(* IEC 61131-3 sources: GenAI/codesys_service/bank/mutants, 40 files *)

(* ---- E01_confirm_level.st ---- *)
FUNCTION_BLOCK E01_Filling
VAR_INPUT
    bottleSensor : BOOL;
    cleaningConfirmButton : BOOL;
    fillingConfirmButton : BOOL;
    cappingConfirmButton : BOOL;
    packingConfirmButton : BOOL;
    finishedButton : BOOL;
END_VAR
VAR_OUTPUT
    Pump_Motor : BOOL;
    Filling_Valve : BOOL;
    Capping_Machine : BOOL;
    Packing_Machine : BOOL;
    Completion_Light : BOOL;
END_VAR
VAR
    step : INT;      (* 0=idle 1=cleaning 2=filling 3=capping 4=packing 5=done *)
    prevBottle : BOOL;
    prevCleaning : BOOL;
    prevFilling : BOOL;
    prevCapping : BOOL;
    prevPacking : BOOL;
    prevFinished : BOOL;
END_VAR

(* step transitions on rising edges *)
IF step = 0 AND bottleSensor AND NOT prevBottle THEN
    step := 1;
END_IF;
IF step = 1 AND cleaningConfirmButton THEN
    step := 2;
END_IF;
IF step = 2 AND fillingConfirmButton THEN
    step := 3;
END_IF;
IF step = 3 AND cappingConfirmButton THEN
    step := 4;
END_IF;
IF step = 4 AND packingConfirmButton THEN
    step := 5;
END_IF;
IF step = 5 AND finishedButton AND NOT prevFinished THEN
    step := 0;
END_IF;

(* outputs by step *)
Pump_Motor := (step = 1);
Filling_Valve := (step = 2);
Capping_Machine := (step = 3);
Packing_Machine := (step = 4);
Completion_Light := (step = 5);

prevBottle := bottleSensor;
prevCleaning := cleaningConfirmButton;
prevFilling := fillingConfirmButton;
prevCapping := cappingConfirmButton;
prevPacking := packingConfirmButton;
prevFinished := finishedButton;

(* ---- E01_no_reset.st ---- *)
FUNCTION_BLOCK E01_Filling
VAR_INPUT
    bottleSensor : BOOL;
    cleaningConfirmButton : BOOL;
    fillingConfirmButton : BOOL;
    cappingConfirmButton : BOOL;
    packingConfirmButton : BOOL;
    finishedButton : BOOL;
END_VAR
VAR_OUTPUT
    Pump_Motor : BOOL;
    Filling_Valve : BOOL;
    Capping_Machine : BOOL;
    Packing_Machine : BOOL;
    Completion_Light : BOOL;
END_VAR
VAR
    step : INT;      (* 0=idle 1=cleaning 2=filling 3=capping 4=packing 5=done *)
    prevBottle : BOOL;
    prevCleaning : BOOL;
    prevFilling : BOOL;
    prevCapping : BOOL;
    prevPacking : BOOL;
    prevFinished : BOOL;
END_VAR

(* step transitions on rising edges *)
IF step = 0 AND bottleSensor AND NOT prevBottle THEN
    step := 1;
END_IF;
IF step = 1 AND cleaningConfirmButton AND NOT prevCleaning THEN
    step := 2;
END_IF;
IF step = 2 AND fillingConfirmButton AND NOT prevFilling THEN
    step := 3;
END_IF;
IF step = 3 AND cappingConfirmButton AND NOT prevCapping THEN
    step := 4;
END_IF;
IF step = 4 AND packingConfirmButton AND NOT prevPacking THEN
    step := 5;
END_IF;
(* bug: finished never resets *)

(* outputs by step *)
Pump_Motor := (step = 1);
Filling_Valve := (step = 2);
Capping_Machine := (step = 3);
Packing_Machine := (step = 4);
Completion_Light := (step = 5);

prevBottle := bottleSensor;
prevCleaning := cleaningConfirmButton;
prevFilling := fillingConfirmButton;
prevCapping := cappingConfirmButton;
prevPacking := packingConfirmButton;
prevFinished := finishedButton;

(* ---- E02_no_prev_update.st ---- *)
(* Q02 Dual-Word Edge Detection - reference solution *)
FUNCTION_BLOCK FB_Q02
VAR_INPUT
    value : DWORD;
END_VAR
VAR_OUTPUT
    hasChanged      : BOOL;
    hasRisingEdges  : BOOL;
    risingBits      : DWORD;
    noOfRisingBits  : USINT;
    hasFallingEdges : BOOL;
    fallingBits     : DWORD;
    noOfFallingBits : USINT;
END_VAR
VAR
    prev : DWORD;
    i    : INT;
    m    : DWORD;
END_VAR

risingBits  := value AND NOT prev;
fallingBits := prev AND NOT value;
hasChanged  := value <> prev;
hasRisingEdges  := risingBits <> 0;
hasFallingEdges := fallingBits <> 0;

noOfRisingBits  := 0;
noOfFallingBits := 0;
FOR i := 0 TO 31 DO
    m := SHL(DWORD#1, i);
    IF (risingBits AND m) <> 0 THEN
        noOfRisingBits := noOfRisingBits + 1;
    END_IF;
    IF (fallingBits AND m) <> 0 THEN
        noOfFallingBits := noOfFallingBits + 1;
    END_IF;
END_FOR;

(* prev not updated *)

(* ---- E02_rising_wrong.st ---- *)
(* Q02 Dual-Word Edge Detection - reference solution *)
FUNCTION_BLOCK FB_Q02
VAR_INPUT
    value : DWORD;
END_VAR
VAR_OUTPUT
    hasChanged      : BOOL;
    hasRisingEdges  : BOOL;
    risingBits      : DWORD;
    noOfRisingBits  : USINT;
    hasFallingEdges : BOOL;
    fallingBits     : DWORD;
    noOfFallingBits : USINT;
END_VAR
VAR
    prev : DWORD;
    i    : INT;
    m    : DWORD;
END_VAR

risingBits  := value;
fallingBits := prev AND NOT value;
hasChanged  := value <> prev;
hasRisingEdges  := risingBits <> 0;
hasFallingEdges := fallingBits <> 0;

noOfRisingBits  := 0;
noOfFallingBits := 0;
FOR i := 0 TO 31 DO
    m := SHL(DWORD#1, i);
    IF (risingBits AND m) <> 0 THEN
        noOfRisingBits := noOfRisingBits + 1;
    END_IF;
    IF (fallingBits AND m) <> 0 THEN
        noOfFallingBits := noOfFallingBits + 1;
    END_IF;
END_FOR;

prev := value;

(* ---- E03_no_hysteresis.st ---- *)
FUNCTION_BLOCK E03_Hysteresis
VAR_INPUT
    Value : REAL;
    hiLevel : REAL;
    loLevel : REAL;
    hystWindow : REAL;
END_VAR
VAR_OUTPUT
    hiAlarm : BOOL;
    loAlarm : BOOL;
    error : BOOL;
    status : WORD;
END_VAR

IF loLevel >= hiLevel THEN
    error := TRUE;
    status := 16#8001;
    hiAlarm := FALSE;
    loAlarm := FALSE;
ELSIF hystWindow >= (hiLevel - loLevel) THEN
    error := TRUE;
    status := 16#8002;
    hiAlarm := FALSE;
    loAlarm := FALSE;
ELSE
    error := FALSE;
    status := 16#0000;
    (* high alarm with hysteresis *)
    IF hiAlarm THEN
        IF Value < hiLevel THEN
            hiAlarm := FALSE;
        END_IF;
    ELSE
        IF Value > hiLevel THEN
            hiAlarm := TRUE;
        END_IF;
    END_IF;
    (* low alarm with hysteresis *)
    IF loAlarm THEN
        IF Value > (loLevel + hystWindow) THEN
            loAlarm := FALSE;
        END_IF;
    ELSE
        IF Value < loLevel THEN
            loAlarm := TRUE;
        END_IF;
    END_IF;
END_IF;

(* ---- E03_no_window_check.st ---- *)
FUNCTION_BLOCK E03_Hysteresis
VAR_INPUT
    Value : REAL;
    hiLevel : REAL;
    loLevel : REAL;
    hystWindow : REAL;
END_VAR
VAR_OUTPUT
    hiAlarm : BOOL;
    loAlarm : BOOL;
    error : BOOL;
    status : WORD;
END_VAR

IF loLevel >= hiLevel THEN
    error := TRUE;
    status := 16#8001;
    hiAlarm := FALSE;
    loAlarm := FALSE;
ELSIF FALSE THEN
    error := TRUE;
    status := 16#8002;
    hiAlarm := FALSE;
    loAlarm := FALSE;
ELSE
    error := FALSE;
    status := 16#0000;
    (* high alarm with hysteresis *)
    IF hiAlarm THEN
        IF Value < (hiLevel - hystWindow) THEN
            hiAlarm := FALSE;
        END_IF;
    ELSE
        IF Value > hiLevel THEN
            hiAlarm := TRUE;
        END_IF;
    END_IF;
    (* low alarm with hysteresis *)
    IF loAlarm THEN
        IF Value > (loLevel + hystWindow) THEN
            loAlarm := FALSE;
        END_IF;
    ELSE
        IF Value < loLevel THEN
            loAlarm := TRUE;
        END_IF;
    END_IF;
END_IF;

(* ---- E04_acc_always.st ---- *)
(* Q04 Jam Pump Debouncing and Runtime Maintenance - reference solution
   Unit convention: TIME inputs in ms, LTIME output in ns (IEC 61131-3). *)
FUNCTION_BLOCK FB_Q04
VAR_INPUT
    VISCOSITY_OK    : BOOL;
    PASTE_E_STOP_NC : BOOL;
    DebounceTime    : TIME;
    CycleTime       : TIME;
END_VAR
VAR_OUTPUT
    VFD_RUN          : BOOL;
    PUMP_MAINT_DUE   : BOOL;
    PUMP_RUNTIME_ACC : LTIME;
END_VAR
VAR
    debAcc  : UDINT;   (* ms *)
    accNs   : ULINT;   (* ns *)
END_VAR

IF NOT PASTE_E_STOP_NC THEN
    VFD_RUN := FALSE;
    debAcc := 0;
ELSE
    IF VISCOSITY_OK THEN
        debAcc := debAcc + TIME_TO_UDINT(CycleTime);
    ELSE
        debAcc := 0;
    END_IF;
    VFD_RUN := VISCOSITY_OK AND debAcc >= TIME_TO_UDINT(DebounceTime);
END_IF;

IF TRUE THEN
    accNs := accNs + UDINT_TO_ULINT(TIME_TO_UDINT(CycleTime)) * 1000000;
    PUMP_RUNTIME_ACC := ULINT_TO_LTIME(accNs);
END_IF;

IF accNs >= 1800000000000000 THEN
    PUMP_MAINT_DUE := TRUE;
END_IF;

(* ---- E04_no_debounce.st ---- *)
(* Q04 Jam Pump Debouncing and Runtime Maintenance - reference solution
   Unit convention: TIME inputs in ms, LTIME output in ns (IEC 61131-3). *)
FUNCTION_BLOCK FB_Q04
VAR_INPUT
    VISCOSITY_OK    : BOOL;
    PASTE_E_STOP_NC : BOOL;
    DebounceTime    : TIME;
    CycleTime       : TIME;
END_VAR
VAR_OUTPUT
    VFD_RUN          : BOOL;
    PUMP_MAINT_DUE   : BOOL;
    PUMP_RUNTIME_ACC : LTIME;
END_VAR
VAR
    debAcc  : UDINT;   (* ms *)
    accNs   : ULINT;   (* ns *)
END_VAR

IF NOT PASTE_E_STOP_NC THEN
    VFD_RUN := FALSE;
    debAcc := 0;
ELSE
    IF VISCOSITY_OK THEN
        debAcc := debAcc + TIME_TO_UDINT(CycleTime);
    ELSE
        debAcc := 0;
    END_IF;
    VFD_RUN := VISCOSITY_OK;
END_IF;

IF VFD_RUN THEN
    accNs := accNs + UDINT_TO_ULINT(TIME_TO_UDINT(CycleTime)) * 1000000;
    PUMP_RUNTIME_ACC := ULINT_TO_LTIME(accNs);
END_IF;

IF accNs >= 1800000000000000 THEN
    PUMP_MAINT_DUE := TRUE;
END_IF;

(* ---- E05_no_estop.st ---- *)
(* Q05 Weld Gap Alarm and Startup Inhibition - reference solution *)
FUNCTION_BLOCK FB_Q05
VAR_INPUT
    Gap_Exceeded   : BOOL;
    Weld_E_Stop_NC : BOOL;
    DebounceTime   : TIME;
END_VAR
VAR_OUTPUT
    Operator_Alert        : BOOL;
    Weld_Soft_Start_Active: BOOL;
END_VAR
VAR
    initTimer : TON;
    debTimer  : TON;
    initDone  : BOOL;
END_VAR

initTimer(IN := Weld_E_Stop_NC AND NOT initDone, PT := T#5S);
IF initTimer.Q THEN
    initDone := TRUE;
END_IF;

IF FALSE THEN
    Operator_Alert := FALSE;
    Weld_Soft_Start_Active := FALSE;
    debTimer(IN := FALSE, PT := DebounceTime);
ELSIF NOT initDone THEN
    Operator_Alert := FALSE;
    Weld_Soft_Start_Active := TRUE;
    debTimer(IN := FALSE, PT := DebounceTime);
ELSE
    Weld_Soft_Start_Active := FALSE;
    debTimer(IN := Gap_Exceeded, PT := DebounceTime);
    Operator_Alert := debTimer.Q;
END_IF;

(* ---- E05_no_inhibit.st ---- *)
(* Q05 Weld Gap Alarm and Startup Inhibition - reference solution *)
FUNCTION_BLOCK FB_Q05
VAR_INPUT
    Gap_Exceeded   : BOOL;
    Weld_E_Stop_NC : BOOL;
    DebounceTime   : TIME;
END_VAR
VAR_OUTPUT
    Operator_Alert        : BOOL;
    Weld_Soft_Start_Active: BOOL;
END_VAR
VAR
    initTimer : TON;
    debTimer  : TON;
    initDone  : BOOL;
END_VAR

initTimer(IN := Weld_E_Stop_NC AND NOT initDone, PT := T#5S);
IF initTimer.Q THEN
    initDone := TRUE;
END_IF;

IF NOT Weld_E_Stop_NC THEN
    Operator_Alert := FALSE;
    Weld_Soft_Start_Active := FALSE;
    debTimer(IN := FALSE, PT := DebounceTime);
ELSIF FALSE THEN
    Operator_Alert := FALSE;
    Weld_Soft_Start_Active := TRUE;
    debTimer(IN := FALSE, PT := DebounceTime);
ELSE
    Weld_Soft_Start_Active := FALSE;
    debTimer(IN := Gap_Exceeded, PT := DebounceTime);
    Operator_Alert := debTimer.Q;
END_IF;

(* ---- E06_count_level.st ---- *)
(* Q06 Aeration Blower Delayed Start - reference solution *)
FUNCTION_BLOCK FB_Q06
VAR_INPUT
    DO_LOW               : BOOL;
    AERATION_E_STOP_NC   : BOOL;
END_VAR
VAR_OUTPUT
    BLOWER_RUN                  : BOOL;
    AERATION_BLOWER_CYCLE_COUNT : UINT;
END_VAR
VAR
    startTimer : TON;
    prevRun    : BOOL;
END_VAR

startTimer(IN := DO_LOW AND AERATION_E_STOP_NC, PT := T#5S);
BLOWER_RUN := startTimer.Q;

IF BLOWER_RUN THEN
    AERATION_BLOWER_CYCLE_COUNT := AERATION_BLOWER_CYCLE_COUNT + 1;
END_IF;
prevRun := BLOWER_RUN;

(* ---- E06_no_delay.st ---- *)
(* Q06 Aeration Blower Delayed Start - reference solution *)
FUNCTION_BLOCK FB_Q06
VAR_INPUT
    DO_LOW               : BOOL;
    AERATION_E_STOP_NC   : BOOL;
END_VAR
VAR_OUTPUT
    BLOWER_RUN                  : BOOL;
    AERATION_BLOWER_CYCLE_COUNT : UINT;
END_VAR
VAR
    startTimer : TON;
    prevRun    : BOOL;
END_VAR

startTimer(IN := DO_LOW AND AERATION_E_STOP_NC, PT := T#5S);
BLOWER_RUN := DO_LOW AND AERATION_E_STOP_NC;

IF BLOWER_RUN AND NOT prevRun THEN
    AERATION_BLOWER_CYCLE_COUNT := AERATION_BLOWER_CYCLE_COUNT + 1;
END_IF;
prevRun := BLOWER_RUN;

(* ---- H01_estop_keeps_step.st ---- *)
FUNCTION_BLOCK H01_Proportion
VAR_INPUT
    estop : BOOL;
    opeMode : BOOL;
    valveAStart : BOOL;
    valveBStart : BOOL;
    valveCStart : BOOL;
    valveDStart : BOOL;
    mixMotorStart : BOOL;
    autoStart : BOOL;
    processMode : BOOL;
    levelSensor : INT;
    mixMotorComplete : BOOL;
END_VAR
VAR_OUTPUT
    valveARun : BOOL;
    valveBRun : BOOL;
    valveCRun : BOOL;
    valveDRun : BOOL;
    mixMotorRun : BOOL;
END_VAR
VAR
    step : INT;  (* 0=idle 1=fillA 2=fillB 3=fillC 4=mixing 5=done *)
    prevAuto : BOOL;
    prevVA : BOOL;
    prevVB : BOOL;
    prevVC : BOOL;
    prevVD : BOOL;
    prevMix : BOOL;
END_VAR

IF NOT estop THEN
    (* emergency stop: everything off, sequence aborted *)
    valveARun := FALSE;
    valveBRun := FALSE;
    valveCRun := FALSE;
    valveDRun := FALSE;
    mixMotorRun := FALSE;
    (* bug: step is kept across the e-stop *)
ELSIF NOT opeMode THEN
    (* manual mode: each button toggles its device on a rising edge *)
    IF valveAStart AND NOT prevVA THEN
        valveARun := NOT valveARun;
    END_IF;
    IF valveBStart AND NOT prevVB THEN
        valveBRun := NOT valveBRun;
    END_IF;
    IF valveCStart AND NOT prevVC THEN
        valveCRun := NOT valveCRun;
    END_IF;
    IF valveDStart AND NOT prevVD THEN
        valveDRun := NOT valveDRun;
    END_IF;
    IF mixMotorStart AND NOT prevMix THEN
        mixMotorRun := NOT mixMotorRun;
    END_IF;
    step := 0;
ELSE
    (* automatic mode state machine *)
    valveCRun := FALSE;
    mixMotorRun := FALSE;
    IF step = 0 THEN
        valveARun := FALSE;
        valveBRun := FALSE;
        valveDRun := FALSE;
        IF autoStart AND NOT prevAuto THEN
            valveARun := TRUE;
            step := 1;
        END_IF;
    ELSIF step = 1 THEN
        valveARun := TRUE;
        IF levelSensor >= 50 THEN
            valveARun := FALSE;
            valveBRun := TRUE;
            step := 2;
        END_IF;
    ELSIF step = 2 THEN
        valveBRun := TRUE;
        IF levelSensor >= 80 THEN
            valveBRun := FALSE;
            IF processMode THEN
                valveCRun := TRUE;
                step := 3;
            ELSE
                mixMotorRun := TRUE;
                step := 4;
            END_IF;
        END_IF;
    ELSIF step = 3 THEN
        valveCRun := TRUE;
        IF levelSensor >= 100 THEN
            valveCRun := FALSE;
            mixMotorRun := TRUE;
            step := 4;
        END_IF;
    ELSIF step = 4 THEN
        mixMotorRun := TRUE;
        IF mixMotorComplete THEN
            mixMotorRun := FALSE;
            valveDRun := TRUE;
            step := 5;
        END_IF;
    ELSE
        (* step 5: process finished, valve D stays open *)
        valveDRun := TRUE;
    END_IF;
END_IF;

prevAuto := autoStart;
prevVA := valveAStart;
prevVB := valveBStart;
prevVC := valveCStart;
prevVD := valveDStart;
prevMix := mixMotorStart;

(* ---- H01_wrong_level.st ---- *)
FUNCTION_BLOCK H01_Proportion
VAR_INPUT
    estop : BOOL;
    opeMode : BOOL;
    valveAStart : BOOL;
    valveBStart : BOOL;
    valveCStart : BOOL;
    valveDStart : BOOL;
    mixMotorStart : BOOL;
    autoStart : BOOL;
    processMode : BOOL;
    levelSensor : INT;
    mixMotorComplete : BOOL;
END_VAR
VAR_OUTPUT
    valveARun : BOOL;
    valveBRun : BOOL;
    valveCRun : BOOL;
    valveDRun : BOOL;
    mixMotorRun : BOOL;
END_VAR
VAR
    step : INT;  (* 0=idle 1=fillA 2=fillB 3=fillC 4=mixing 5=done *)
    prevAuto : BOOL;
    prevVA : BOOL;
    prevVB : BOOL;
    prevVC : BOOL;
    prevVD : BOOL;
    prevMix : BOOL;
END_VAR

IF NOT estop THEN
    (* emergency stop: everything off, sequence aborted *)
    valveARun := FALSE;
    valveBRun := FALSE;
    valveCRun := FALSE;
    valveDRun := FALSE;
    mixMotorRun := FALSE;
    step := 0;
ELSIF NOT opeMode THEN
    (* manual mode: each button toggles its device on a rising edge *)
    IF valveAStart AND NOT prevVA THEN
        valveARun := NOT valveARun;
    END_IF;
    IF valveBStart AND NOT prevVB THEN
        valveBRun := NOT valveBRun;
    END_IF;
    IF valveCStart AND NOT prevVC THEN
        valveCRun := NOT valveCRun;
    END_IF;
    IF valveDStart AND NOT prevVD THEN
        valveDRun := NOT valveDRun;
    END_IF;
    IF mixMotorStart AND NOT prevMix THEN
        mixMotorRun := NOT mixMotorRun;
    END_IF;
    step := 0;
ELSE
    (* automatic mode state machine *)
    valveCRun := FALSE;
    mixMotorRun := FALSE;
    IF step = 0 THEN
        valveARun := FALSE;
        valveBRun := FALSE;
        valveDRun := FALSE;
        IF autoStart AND NOT prevAuto THEN
            valveARun := TRUE;
            step := 1;
        END_IF;
    ELSIF step = 1 THEN
        valveARun := TRUE;
        IF levelSensor >= 60 THEN
            valveARun := FALSE;
            valveBRun := TRUE;
            step := 2;
        END_IF;
    ELSIF step = 2 THEN
        valveBRun := TRUE;
        IF levelSensor >= 80 THEN
            valveBRun := FALSE;
            IF processMode THEN
                valveCRun := TRUE;
                step := 3;
            ELSE
                mixMotorRun := TRUE;
                step := 4;
            END_IF;
        END_IF;
    ELSIF step = 3 THEN
        valveCRun := TRUE;
        IF levelSensor >= 100 THEN
            valveCRun := FALSE;
            mixMotorRun := TRUE;
            step := 4;
        END_IF;
    ELSIF step = 4 THEN
        mixMotorRun := TRUE;
        IF mixMotorComplete THEN
            mixMotorRun := FALSE;
            valveDRun := TRUE;
            step := 5;
        END_IF;
    ELSE
        (* step 5: process finished, valve D stays open *)
        valveDRun := TRUE;
    END_IF;
END_IF;

prevAuto := autoStart;
prevVA := valveAStart;
prevVB := valveBStart;
prevVC := valveCStart;
prevVD := valveDStart;
prevMix := mixMotorStart;

(* ---- H02_always_right.st ---- *)
(* Q16 Flexible Processing Control - reference solution *)
FUNCTION_BLOCK FB_Q16
VAR_INPUT
    processLength   : USINT;
    sensor1         : BOOL;
    sensor2         : BOOL;
    sensor3         : BOOL;
    sensor4         : BOOL;
    sensor5         : BOOL;
    station1Start   : BOOL;
    station2Complete: BOOL;
    station3Complete: BOOL;
    station4Complete: BOOL;
    processSequence : ARRAY[1..8] OF USINT;
END_VAR
VAR_OUTPUT
    conveyorLeft  : BOOL;
    conveyorRight : BOOL;
END_VAR
VAR
    idx     : USINT;      (* active entry, 0 = not started *)
    cur     : USINT;      (* station the product is at, 0 = in transit *)
    target  : USINT;
    moving  : BOOL;
    atTarget: BOOL;
    done    : BOOL;
END_VAR

conveyorLeft := FALSE;
conveyorRight := FALSE;

(* current station from the sensors *)
cur := 0;
IF sensor1 THEN cur := 1; END_IF;
IF sensor2 THEN cur := 2; END_IF;
IF sensor3 THEN cur := 3; END_IF;
IF sensor4 THEN cur := 4; END_IF;
IF sensor5 THEN cur := 5; END_IF;

IF idx = 0 THEN
    IF sensor1 AND station1Start THEN
        idx := 1;
        moving := TRUE;
    END_IF;
ELSE
    target := processSequence[idx];
    atTarget := (cur = target);

    IF moving AND atTarget THEN
        moving := FALSE;                     (* arrived: stop *)
    END_IF;

    IF NOT moving AND atTarget THEN
        done := FALSE;
        IF target = 2 THEN
            done := station2Complete;
        ELSIF target = 3 THEN
            done := station3Complete;
        ELSIF target = 4 THEN
            done := station4Complete;
        END_IF;
        IF done AND idx < processLength THEN
            idx := idx + 1;
            moving := TRUE;
        END_IF;
    END_IF;

    IF moving THEN
        target := processSequence[idx];
        IF cur = 0 THEN
            (* in transit: keep the previous direction *)
            conveyorRight := conveyorRight OR NOT conveyorLeft;
        END_IF;
        IF target > cur AND cur > 0 THEN
            conveyorRight := TRUE;
        ELSIF FALSE THEN
            conveyorLeft := TRUE;
        END_IF;
    END_IF;
END_IF;

(* ---- H02_no_wait.st ---- *)
(* Q16 Flexible Processing Control - reference solution *)
FUNCTION_BLOCK FB_Q16
VAR_INPUT
    processLength   : USINT;
    sensor1         : BOOL;
    sensor2         : BOOL;
    sensor3         : BOOL;
    sensor4         : BOOL;
    sensor5         : BOOL;
    station1Start   : BOOL;
    station2Complete: BOOL;
    station3Complete: BOOL;
    station4Complete: BOOL;
    processSequence : ARRAY[1..8] OF USINT;
END_VAR
VAR_OUTPUT
    conveyorLeft  : BOOL;
    conveyorRight : BOOL;
END_VAR
VAR
    idx     : USINT;      (* active entry, 0 = not started *)
    cur     : USINT;      (* station the product is at, 0 = in transit *)
    target  : USINT;
    moving  : BOOL;
    atTarget: BOOL;
    done    : BOOL;
END_VAR

conveyorLeft := FALSE;
conveyorRight := FALSE;

(* current station from the sensors *)
cur := 0;
IF sensor1 THEN cur := 1; END_IF;
IF sensor2 THEN cur := 2; END_IF;
IF sensor3 THEN cur := 3; END_IF;
IF sensor4 THEN cur := 4; END_IF;
IF sensor5 THEN cur := 5; END_IF;

IF idx = 0 THEN
    IF sensor1 AND station1Start THEN
        idx := 1;
        moving := TRUE;
    END_IF;
ELSE
    target := processSequence[idx];
    atTarget := (cur = target);

    IF moving AND atTarget THEN
        moving := FALSE;                     (* arrived: stop *)
    END_IF;

    IF NOT moving AND atTarget THEN
        done := FALSE;
        IF target = 2 THEN
            done := station2Complete;
        ELSIF target = 3 THEN
            done := station3Complete;
        ELSIF target = 4 THEN
            done := station4Complete;
        END_IF;
        IF idx < processLength THEN
            idx := idx + 1;
            moving := TRUE;
        END_IF;
    END_IF;

    IF moving THEN
        target := processSequence[idx];
        IF cur = 0 THEN
            (* in transit: keep the previous direction *)
            conveyorRight := conveyorRight OR NOT conveyorLeft;
        END_IF;
        IF target > cur AND cur > 0 THEN
            conveyorRight := TRUE;
        ELSIF target < cur AND cur > 0 THEN
            conveyorLeft := TRUE;
        END_IF;
    END_IF;
END_IF;

(* ---- H03_delete_wrong_code.st ---- *)
TYPE ST_Recipe :
STRUCT
    recipeID              : INT;
    ingredientType        : INT;
    ingredientRatio       : REAL;
    productionTemperature : REAL;
END_STRUCT
END_TYPE

(* Q17 Recipe Management System - reference solution *)
FUNCTION_BLOCK FB_Q17
VAR_INPUT
    addRecipe    : BOOL;
    deleteRecipe : BOOL;
    modifyRecipe : BOOL;
    queryRecipe  : BOOL;
    recipeIn     : ST_Recipe;
END_VAR
VAR_OUTPUT
    recipeAdded       : BOOL;
    recipeDeleted     : BOOL;
    recipeModified    : BOOL;
    recipeQueryResult : ST_Recipe;
    error             : BOOL;
    status            : WORD;
END_VAR
VAR_IN_OUT
    recipe : ARRAY[1..10] OF ST_Recipe;
END_VAR
VAR
    i    : INT;
    slot : INT;
    free : INT;
END_VAR

recipeAdded := FALSE;
recipeDeleted := FALSE;
recipeModified := FALSE;
error := FALSE;
status := 16#0000;

slot := 0;
free := 0;
FOR i := 10 TO 1 BY -1 DO
    IF recipe[i].recipeID = recipeIn.recipeID THEN
        slot := i;
    END_IF;
    IF recipe[i].recipeID = 0 THEN
        free := i;
    END_IF;
END_FOR;

IF queryRecipe THEN
    IF slot = 0 THEN
        error := TRUE;
        status := 16#8001;
    ELSE
        recipeQueryResult := recipe[slot];
    END_IF;
ELSIF addRecipe THEN
    IF slot <> 0 THEN
        error := TRUE;
        status := 16#8002;
    ELSIF free = 0 THEN
        error := TRUE;
        status := 16#8003;
    ELSE
        recipe[free] := recipeIn;
        recipeAdded := TRUE;
    END_IF;
ELSIF deleteRecipe THEN
    IF slot = 0 THEN
        error := TRUE;
        status := 16#8001;
    ELSE
        recipe[slot].recipeID := 0;
        recipeDeleted := TRUE;
    END_IF;
ELSIF modifyRecipe THEN
    IF slot = 0 THEN
        error := TRUE;
        status := 16#8005;
    ELSE
        recipe[slot] := recipeIn;
        recipeModified := TRUE;
    END_IF;
END_IF;

(* ---- H03_no_dup_check.st ---- *)
TYPE ST_Recipe :
STRUCT
    recipeID              : INT;
    ingredientType        : INT;
    ingredientRatio       : REAL;
    productionTemperature : REAL;
END_STRUCT
END_TYPE

(* Q17 Recipe Management System - reference solution *)
FUNCTION_BLOCK FB_Q17
VAR_INPUT
    addRecipe    : BOOL;
    deleteRecipe : BOOL;
    modifyRecipe : BOOL;
    queryRecipe  : BOOL;
    recipeIn     : ST_Recipe;
END_VAR
VAR_OUTPUT
    recipeAdded       : BOOL;
    recipeDeleted     : BOOL;
    recipeModified    : BOOL;
    recipeQueryResult : ST_Recipe;
    error             : BOOL;
    status            : WORD;
END_VAR
VAR_IN_OUT
    recipe : ARRAY[1..10] OF ST_Recipe;
END_VAR
VAR
    i    : INT;
    slot : INT;
    free : INT;
END_VAR

recipeAdded := FALSE;
recipeDeleted := FALSE;
recipeModified := FALSE;
error := FALSE;
status := 16#0000;

slot := 0;
free := 0;
FOR i := 10 TO 1 BY -1 DO
    IF recipe[i].recipeID = recipeIn.recipeID THEN
        slot := i;
    END_IF;
    IF recipe[i].recipeID = 0 THEN
        free := i;
    END_IF;
END_FOR;

IF queryRecipe THEN
    IF slot = 0 THEN
        error := TRUE;
        status := 16#8001;
    ELSE
        recipeQueryResult := recipe[slot];
    END_IF;
ELSIF addRecipe THEN
    IF FALSE THEN
        error := TRUE;
        status := 16#8002;
    ELSIF free = 0 THEN
        error := TRUE;
        status := 16#8003;
    ELSE
        recipe[free] := recipeIn;
        recipeAdded := TRUE;
    END_IF;
ELSIF deleteRecipe THEN
    IF slot = 0 THEN
        error := TRUE;
        status := 16#8004;
    ELSE
        recipe[slot].recipeID := 0;
        recipeDeleted := TRUE;
    END_IF;
ELSIF modifyRecipe THEN
    IF slot = 0 THEN
        error := TRUE;
        status := 16#8005;
    ELSE
        recipe[slot] := recipeIn;
        recipeModified := TRUE;
    END_IF;
END_IF;

(* ---- H04_enq_level.st ---- *)
(* Q18 FIFO Queue - reference solution.
   The interface uses VARIANT in the task; this reference uses a concrete
   INT array so that it can be compiled and tested in the harness. *)
FUNCTION_BLOCK FB_Q18
VAR_INPUT
    enqueue : BOOL;
    dequeue : BOOL;
    reset   : BOOL;
END_VAR
VAR_OUTPUT
    elementCount : DINT;
    status       : WORD;
END_VAR
VAR_IN_OUT
    item   : INT;
    buffer : ARRAY[1..5] OF INT;
END_VAR
VAR
    head : DINT := 1;
    tail : DINT := 1;
    cap  : DINT := 5;
    prevEnq : BOOL;
    prevDeq : BOOL;
    enqEdge : BOOL;
    deqEdge : BOOL;
END_VAR

status := 16#0000;
enqEdge := enqueue;
deqEdge := dequeue AND NOT prevDeq;
prevEnq := enqueue;
prevDeq := dequeue;

IF reset THEN
    head := 1;
    tail := 1;
    elementCount := 0;
ELSIF enqEdge THEN
    IF elementCount >= cap THEN
        status := 16#8002;
    ELSE
        buffer[tail] := item;
        tail := tail + 1;
        IF tail > cap THEN
            tail := 1;
        END_IF;
        elementCount := elementCount + 1;
    END_IF;
ELSIF deqEdge THEN
    IF elementCount <= 0 THEN
        status := 16#8001;
    ELSE
        item := buffer[head];
        head := head + 1;
        IF head > cap THEN
            head := 1;
        END_IF;
        elementCount := elementCount - 1;
    END_IF;
END_IF;

(* ---- H04_no_full_check.st ---- *)
(* Q18 FIFO Queue - reference solution.
   The interface uses VARIANT in the task; this reference uses a concrete
   INT array so that it can be compiled and tested in the harness. *)
FUNCTION_BLOCK FB_Q18
VAR_INPUT
    enqueue : BOOL;
    dequeue : BOOL;
    reset   : BOOL;
END_VAR
VAR_OUTPUT
    elementCount : DINT;
    status       : WORD;
END_VAR
VAR_IN_OUT
    item   : INT;
    buffer : ARRAY[1..5] OF INT;
END_VAR
VAR
    head : DINT := 1;
    tail : DINT := 1;
    cap  : DINT := 5;
    prevEnq : BOOL;
    prevDeq : BOOL;
    enqEdge : BOOL;
    deqEdge : BOOL;
END_VAR

status := 16#0000;
enqEdge := enqueue AND NOT prevEnq;
deqEdge := dequeue AND NOT prevDeq;
prevEnq := enqueue;
prevDeq := dequeue;

IF reset THEN
    head := 1;
    tail := 1;
    elementCount := 0;
ELSIF enqEdge THEN
    IF FALSE THEN
        status := 16#8002;
    ELSE
        buffer[tail] := item;
        tail := tail + 1;
        IF tail > cap THEN
            tail := 1;
        END_IF;
        elementCount := elementCount + 1;
    END_IF;
ELSIF deqEdge THEN
    IF elementCount <= 0 THEN
        status := 16#8001;
    ELSE
        item := buffer[head];
        head := head + 1;
        IF head > cap THEN
            head := 1;
        END_IF;
        elementCount := elementCount - 1;
    END_IF;
END_IF;

(* ---- H05_ignore_limits.st ---- *)
FUNCTION_BLOCK H05_MechArm
VAR_INPUT
    ManualMode : BOOL;
    SingleStepMode : BOOL;
    SingleCycleMode : BOOL;
    ContinuousMode : BOOL;
    EmergencyStop : BOOL;
    Start : BOOL;
    DownButton : BOOL;
    UpButton : BOOL;
    LeftButton : BOOL;
    RightButton : BOOL;
    GripButton : BOOL;
    ReleaseButton : BOOL;
    DownLimitSwitch : BOOL;
    UpLimitSwitch : BOOL;
    LeftLimitSwitch : BOOL;
    RightLimitSwitch : BOOL;
    GripLimitSwitch : BOOL;
    ReleaseLimitSwitch : BOOL;
END_VAR
VAR_OUTPUT
    MoveDown : BOOL;
    MoveUp : BOOL;
    MoveLeft : BOOL;
    MoveRight : BOOL;
    ActivateGrip : BOOL;
    ActivateRelease : BOOL;
END_VAR
VAR
    step : INT := 0;   (* 0 idle, then 1..8 = the 8-action cycle *)
    prevStart : BOOL;
    running : BOOL;
END_VAR

MoveDown := FALSE;
MoveUp := FALSE;
MoveLeft := FALSE;
MoveRight := FALSE;
ActivateGrip := FALSE;
ActivateRelease := FALSE;

IF NOT EmergencyStop THEN
    (* emergency stop: all actions off, sequence aborted *)
    step := 0;
    running := FALSE;
ELSIF ManualMode THEN
    (* manual: buttons drive actions, limited by position switches *)
    MoveDown := DownButton;
    MoveUp := UpButton;
    MoveLeft := LeftButton;
    MoveRight := RightButton;
    ActivateGrip := GripButton AND NOT GripLimitSwitch;
    ActivateRelease := ReleaseButton AND NOT ReleaseLimitSwitch;
    step := 0;
    running := FALSE;
ELSIF SingleStepMode THEN
    (* single step: each start press advances one action *)
    IF Start AND NOT prevStart AND NOT running THEN
        IF step = 0 THEN
            step := 1;
        END_IF;
    END_IF;
    IF step > 0 THEN
        running := TRUE;
    END_IF;
ELSE
    (* single cycle / continuous: run through the cycle automatically *)
    IF (Start AND NOT prevStart) AND (step = 0) THEN
        step := 1;
    END_IF;
    IF step > 0 THEN
        running := TRUE;
    END_IF;
END_IF;

IF running AND EmergencyStop THEN
    (* action execution by step; each step stops on its completion feedback *)
    IF step = 1 THEN
        MoveDown := NOT DownLimitSwitch;
        IF DownLimitSwitch THEN step := 2; END_IF;
    ELSIF step = 2 THEN
        ActivateGrip := NOT GripLimitSwitch;
        IF GripLimitSwitch THEN step := 3; END_IF;
    ELSIF step = 3 THEN
        MoveUp := NOT UpLimitSwitch;
        IF UpLimitSwitch THEN step := 4; END_IF;
    ELSIF step = 4 THEN
        MoveRight := NOT RightLimitSwitch;
        IF RightLimitSwitch THEN step := 5; END_IF;
    ELSIF step = 5 THEN
        MoveDown := NOT DownLimitSwitch;
        IF DownLimitSwitch THEN step := 6; END_IF;
    ELSIF step = 6 THEN
        ActivateRelease := NOT ReleaseLimitSwitch;
        IF ReleaseLimitSwitch THEN step := 7; END_IF;
    ELSIF step = 7 THEN
        MoveUp := NOT UpLimitSwitch;
        IF UpLimitSwitch THEN step := 8; END_IF;
    ELSIF step = 8 THEN
        MoveLeft := NOT LeftLimitSwitch;
        IF LeftLimitSwitch THEN
            (* cycle complete: single cycle stops, continuous restarts *)
            IF ContinuousMode THEN
                step := 1;
            ELSE
                step := 0;
                running := FALSE;
            END_IF;
        END_IF;
    ELSE
        running := FALSE;
    END_IF;

    (* single step pauses between actions after completing one *)
    IF SingleStepMode AND (step > 1) THEN
        (* stop execution after the current action finishes:
           handled implicitly on the next invocation *)
        running := FALSE;
        step := step;  (* hold position, wait for next start *)
    END_IF;
END_IF;

prevStart := Start;

(* ---- H05_no_continuous_restart.st ---- *)
FUNCTION_BLOCK H05_MechArm
VAR_INPUT
    ManualMode : BOOL;
    SingleStepMode : BOOL;
    SingleCycleMode : BOOL;
    ContinuousMode : BOOL;
    EmergencyStop : BOOL;
    Start : BOOL;
    DownButton : BOOL;
    UpButton : BOOL;
    LeftButton : BOOL;
    RightButton : BOOL;
    GripButton : BOOL;
    ReleaseButton : BOOL;
    DownLimitSwitch : BOOL;
    UpLimitSwitch : BOOL;
    LeftLimitSwitch : BOOL;
    RightLimitSwitch : BOOL;
    GripLimitSwitch : BOOL;
    ReleaseLimitSwitch : BOOL;
END_VAR
VAR_OUTPUT
    MoveDown : BOOL;
    MoveUp : BOOL;
    MoveLeft : BOOL;
    MoveRight : BOOL;
    ActivateGrip : BOOL;
    ActivateRelease : BOOL;
END_VAR
VAR
    step : INT := 0;   (* 0 idle, then 1..8 = the 8-action cycle *)
    prevStart : BOOL;
    running : BOOL;
END_VAR

MoveDown := FALSE;
MoveUp := FALSE;
MoveLeft := FALSE;
MoveRight := FALSE;
ActivateGrip := FALSE;
ActivateRelease := FALSE;

IF NOT EmergencyStop THEN
    (* emergency stop: all actions off, sequence aborted *)
    step := 0;
    running := FALSE;
ELSIF ManualMode THEN
    (* manual: buttons drive actions, limited by position switches *)
    MoveDown := DownButton AND NOT DownLimitSwitch;
    MoveUp := UpButton AND NOT UpLimitSwitch;
    MoveLeft := LeftButton AND NOT LeftLimitSwitch;
    MoveRight := RightButton AND NOT RightLimitSwitch;
    ActivateGrip := GripButton AND NOT GripLimitSwitch;
    ActivateRelease := ReleaseButton AND NOT ReleaseLimitSwitch;
    step := 0;
    running := FALSE;
ELSIF SingleStepMode THEN
    (* single step: each start press advances one action *)
    IF Start AND NOT prevStart AND NOT running THEN
        IF step = 0 THEN
            step := 1;
        END_IF;
    END_IF;
    IF step > 0 THEN
        running := TRUE;
    END_IF;
ELSE
    (* single cycle / continuous: run through the cycle automatically *)
    IF (Start AND NOT prevStart) AND (step = 0) THEN
        step := 1;
    END_IF;
    IF step > 0 THEN
        running := TRUE;
    END_IF;
END_IF;

IF running AND EmergencyStop THEN
    (* action execution by step; each step stops on its completion feedback *)
    IF step = 1 THEN
        MoveDown := NOT DownLimitSwitch;
        IF DownLimitSwitch THEN step := 2; END_IF;
    ELSIF step = 2 THEN
        ActivateGrip := NOT GripLimitSwitch;
        IF GripLimitSwitch THEN step := 3; END_IF;
    ELSIF step = 3 THEN
        MoveUp := NOT UpLimitSwitch;
        IF UpLimitSwitch THEN step := 4; END_IF;
    ELSIF step = 4 THEN
        MoveRight := NOT RightLimitSwitch;
        IF RightLimitSwitch THEN step := 5; END_IF;
    ELSIF step = 5 THEN
        MoveDown := NOT DownLimitSwitch;
        IF DownLimitSwitch THEN step := 6; END_IF;
    ELSIF step = 6 THEN
        ActivateRelease := NOT ReleaseLimitSwitch;
        IF ReleaseLimitSwitch THEN step := 7; END_IF;
    ELSIF step = 7 THEN
        MoveUp := NOT UpLimitSwitch;
        IF UpLimitSwitch THEN step := 8; END_IF;
    ELSIF step = 8 THEN
        MoveLeft := NOT LeftLimitSwitch;
        IF LeftLimitSwitch THEN
            (* cycle complete: single cycle stops, continuous restarts *)
            (* bug: continuous mode does not restart the cycle *)
            step := 0;
            running := FALSE;
        END_IF;
    ELSE
        running := FALSE;
    END_IF;

    (* single step pauses between actions after completing one *)
    IF SingleStepMode AND (step > 1) THEN
        (* stop execution after the current action finishes:
           handled implicitly on the next invocation *)
        running := FALSE;
        step := step;  (* hold position, wait for next start *)
    END_IF;
END_IF;

prevStart := Start;

(* ---- H06_no_upper_limit.st ---- *)
FUNCTION_BLOCK H06_Production
VAR_INPUT
    Mode : BOOL;
    ForwardButton : BOOL;
    ReverseButton : BOOL;
    SensorFeed : BOOL;
    SensorWash : BOOL;
    SensorWeight : BOOL;
    SensorFiring : BOOL;
    SensorOutput : BOOL;
    washComplete : BOOL;
    weightComplete : BOOL;
    weight : REAL;
    firingComplete : BOOL;
END_VAR
VAR_OUTPUT
    MotorForward : BOOL;
    MotorReverse : BOOL;
    kick : BOOL;
    CompletionLight : BOOL;
    firingTemp : REAL;
END_VAR
VAR
    step : INT;  (* 0=feed 1=feed->wash 2=wash wait 3=wash->weight 4=weigh
                    5=weight->(kick|fire) 6=fire wait 7=fire->out 8=done *)
    qualified : BOOL;
    prevWashC : BOOL;
    prevWeightC : BOOL;
    prevFireC : BOOL;
END_VAR

IF NOT Mode THEN
    MotorForward := ForwardButton AND NOT ReverseButton;
    MotorReverse := ReverseButton AND NOT ForwardButton;
    kick := FALSE;
    CompletionLight := FALSE;
    step := 0;
ELSE
    MotorReverse := FALSE;
    IF step = 0 THEN
        MotorForward := FALSE;
        kick := FALSE;
        IF SensorFeed THEN
            step := 1;
        END_IF;
    ELSIF step = 1 THEN
        MotorForward := TRUE;
        IF SensorWash THEN
            MotorForward := FALSE;
            step := 2;
        END_IF;
    ELSIF step = 2 THEN
        MotorForward := FALSE;
        IF washComplete AND NOT prevWashC THEN
            step := 3;
        END_IF;
    ELSIF step = 3 THEN
        MotorForward := TRUE;
        IF SensorWeight THEN
            MotorForward := FALSE;
            step := 4;
        END_IF;
    ELSIF step = 4 THEN
        MotorForward := FALSE;
        IF weightComplete AND NOT prevWeightC THEN
            qualified := (weight >= 100.0);
            IF qualified THEN
                (* 100..200 kg -> 500..550 degrees, linear *)
                firingTemp := 500.0 + (weight - 100.0) * 0.5;
                step := 5;
            ELSE
                kick := TRUE;
                step := 8;
            END_IF;
        END_IF;
    ELSIF step = 5 THEN
        MotorForward := TRUE;
        IF SensorFiring THEN
            MotorForward := FALSE;
            step := 6;
        END_IF;
    ELSIF step = 6 THEN
        MotorForward := FALSE;
        IF firingComplete AND NOT prevFireC THEN
            step := 7;
        END_IF;
    ELSIF step = 7 THEN
        MotorForward := TRUE;
        IF SensorOutput THEN
            MotorForward := FALSE;
            step := 8;
        END_IF;
    ELSE
        (* step 8: finished / rejected *)
        MotorForward := FALSE;
        CompletionLight := SensorOutput;
        IF NOT SensorOutput THEN
            CompletionLight := FALSE;
            kick := FALSE;
            step := 0;
        END_IF;
    END_IF;
END_IF;

prevWashC := washComplete;
prevWeightC := weightComplete;
prevFireC := firingComplete;

(* ---- H06_wrong_temp.st ---- *)
FUNCTION_BLOCK H06_Production
VAR_INPUT
    Mode : BOOL;
    ForwardButton : BOOL;
    ReverseButton : BOOL;
    SensorFeed : BOOL;
    SensorWash : BOOL;
    SensorWeight : BOOL;
    SensorFiring : BOOL;
    SensorOutput : BOOL;
    washComplete : BOOL;
    weightComplete : BOOL;
    weight : REAL;
    firingComplete : BOOL;
END_VAR
VAR_OUTPUT
    MotorForward : BOOL;
    MotorReverse : BOOL;
    kick : BOOL;
    CompletionLight : BOOL;
    firingTemp : REAL;
END_VAR
VAR
    step : INT;  (* 0=feed 1=feed->wash 2=wash wait 3=wash->weight 4=weigh
                    5=weight->(kick|fire) 6=fire wait 7=fire->out 8=done *)
    qualified : BOOL;
    prevWashC : BOOL;
    prevWeightC : BOOL;
    prevFireC : BOOL;
END_VAR

IF NOT Mode THEN
    MotorForward := ForwardButton AND NOT ReverseButton;
    MotorReverse := ReverseButton AND NOT ForwardButton;
    kick := FALSE;
    CompletionLight := FALSE;
    step := 0;
ELSE
    MotorReverse := FALSE;
    IF step = 0 THEN
        MotorForward := FALSE;
        kick := FALSE;
        IF SensorFeed THEN
            step := 1;
        END_IF;
    ELSIF step = 1 THEN
        MotorForward := TRUE;
        IF SensorWash THEN
            MotorForward := FALSE;
            step := 2;
        END_IF;
    ELSIF step = 2 THEN
        MotorForward := FALSE;
        IF washComplete AND NOT prevWashC THEN
            step := 3;
        END_IF;
    ELSIF step = 3 THEN
        MotorForward := TRUE;
        IF SensorWeight THEN
            MotorForward := FALSE;
            step := 4;
        END_IF;
    ELSIF step = 4 THEN
        MotorForward := FALSE;
        IF weightComplete AND NOT prevWeightC THEN
            qualified := (weight >= 100.0) AND (weight <= 200.0);
            IF qualified THEN
                (* 100..200 kg -> 500..550 degrees, linear *)
                firingTemp := 500.0 + (weight - 100.0) * 1.0;
                step := 5;
            ELSE
                kick := TRUE;
                step := 8;
            END_IF;
        END_IF;
    ELSIF step = 5 THEN
        MotorForward := TRUE;
        IF SensorFiring THEN
            MotorForward := FALSE;
            step := 6;
        END_IF;
    ELSIF step = 6 THEN
        MotorForward := FALSE;
        IF firingComplete AND NOT prevFireC THEN
            step := 7;
        END_IF;
    ELSIF step = 7 THEN
        MotorForward := TRUE;
        IF SensorOutput THEN
            MotorForward := FALSE;
            step := 8;
        END_IF;
    ELSE
        (* step 8: finished / rejected *)
        MotorForward := FALSE;
        CompletionLight := SensorOutput;
        IF NOT SensorOutput THEN
            CompletionLight := FALSE;
            kick := FALSE;
            step := 0;
        END_IF;
    END_IF;
END_IF;

prevWashC := washComplete;
prevWeightC := weightComplete;
prevFireC := firingComplete;

(* ---- M01_manual_ignores_sel.st ---- *)
TYPE ST_Pump :
STRUCT
    priority  : INT;
    selection : BOOL;
    RunComd   : BOOL;
END_STRUCT
END_TYPE

(* Q07 Multi-Pump Switching Control System - reference solution *)
FUNCTION_BLOCK FB_Q07
VAR_INPUT
    mode  : BOOL;
    start : BOOL;
    stop  : BOOL;
END_VAR
VAR_IN_OUT
    pumpGroup : ARRAY[1..5] OF ST_Pump;
END_VAR
VAR
    i, j, best, bestIdx, picked : INT;
    chosen : ARRAY[1..5] OF BOOL;
    running : BOOL;
END_VAR

IF stop THEN
    FOR i := 1 TO 5 DO
        pumpGroup[i].RunComd := FALSE;
    END_FOR;
    running := FALSE;
ELSIF start THEN
    running := TRUE;
END_IF;

IF running THEN
    IF NOT mode THEN
        (* manual: run exactly the selected pumps *)
        FOR i := 1 TO 5 DO
            pumpGroup[i].RunComd := TRUE;
        END_FOR;
    ELSE
        (* automatic: three highest priorities run, two stand by *)
        FOR i := 1 TO 5 DO
            chosen[i] := FALSE;
        END_FOR;
        FOR picked := 1 TO 3 DO
            bestIdx := 0;
            FOR j := 1 TO 5 DO
                IF NOT chosen[j] THEN
                    IF bestIdx = 0 THEN
                        bestIdx := j;
                        best := pumpGroup[j].priority;
                    ELSIF pumpGroup[j].priority > best THEN
                        bestIdx := j;
                        best := pumpGroup[j].priority;
                    END_IF;
                END_IF;
            END_FOR;
            IF bestIdx > 0 THEN
                chosen[bestIdx] := TRUE;
            END_IF;
        END_FOR;
        FOR i := 1 TO 5 DO
            pumpGroup[i].RunComd := chosen[i];
        END_FOR;
    END_IF;
END_IF;

(* ---- M01_pick_two.st ---- *)
TYPE ST_Pump :
STRUCT
    priority  : INT;
    selection : BOOL;
    RunComd   : BOOL;
END_STRUCT
END_TYPE

(* Q07 Multi-Pump Switching Control System - reference solution *)
FUNCTION_BLOCK FB_Q07
VAR_INPUT
    mode  : BOOL;
    start : BOOL;
    stop  : BOOL;
END_VAR
VAR_IN_OUT
    pumpGroup : ARRAY[1..5] OF ST_Pump;
END_VAR
VAR
    i, j, best, bestIdx, picked : INT;
    chosen : ARRAY[1..5] OF BOOL;
    running : BOOL;
END_VAR

IF stop THEN
    FOR i := 1 TO 5 DO
        pumpGroup[i].RunComd := FALSE;
    END_FOR;
    running := FALSE;
ELSIF start THEN
    running := TRUE;
END_IF;

IF running THEN
    IF NOT mode THEN
        (* manual: run exactly the selected pumps *)
        FOR i := 1 TO 5 DO
            pumpGroup[i].RunComd := pumpGroup[i].selection;
        END_FOR;
    ELSE
        (* automatic: three highest priorities run, two stand by *)
        FOR i := 1 TO 5 DO
            chosen[i] := FALSE;
        END_FOR;
        FOR picked := 1 TO 2 DO
            bestIdx := 0;
            FOR j := 1 TO 5 DO
                IF NOT chosen[j] THEN
                    IF bestIdx = 0 THEN
                        bestIdx := j;
                        best := pumpGroup[j].priority;
                    ELSIF pumpGroup[j].priority > best THEN
                        bestIdx := j;
                        best := pumpGroup[j].priority;
                    END_IF;
                END_IF;
            END_FOR;
            IF bestIdx > 0 THEN
                chosen[bestIdx] := TRUE;
            END_IF;
        END_FOR;
        FOR i := 1 TO 5 DO
            pumpGroup[i].RunComd := chosen[i];
        END_FOR;
    END_IF;
END_IF;

(* ---- M02_limit_check_off.st ---- *)
TYPE ST_AnalogChannel :
STRUCT
    enable        : BOOL;
    hiLIM         : REAL;
    loLIM         : REAL;
    bipolar       : BOOL;
    measuringMode : INT;
    retVal        : WORD;
    outputValue   : REAL;
END_STRUCT
END_TYPE

(* Q08 Analog Batch Processing - reference solution.
   The task declares ARRAY[*]; this reference fixes the length at 2 so that it
   can be compiled and exercised by the test harness. *)
FUNCTION_BLOCK FB_Q08
VAR_INPUT
    count : DINT;
END_VAR
VAR_IN_OUT
    analogValues : ARRAY[1..2] OF INT;
    channels     : ARRAY[1..2] OF ST_AnalogChannel;
END_VAR
VAR
    i   : DINT;
    raw : REAL;
END_VAR

FOR i := 1 TO 2 DO
    IF i <= count AND channels[i].enable THEN
        IF channels[i].measuringMode < 0 OR channels[i].measuringMode > 2 THEN
            channels[i].retVal := 16#8001;
        ELSIF channels[i].hiLIM < channels[i].loLIM THEN
            channels[i].retVal := 16#8002;
        ELSE
            channels[i].retVal := 16#0000;
            raw := INT_TO_REAL(analogValues[i]);
            IF channels[i].measuringMode = 0 THEN
                IF channels[i].bipolar THEN
                    channels[i].outputValue := channels[i].loLIM
                        + (raw + 27648.0) / 55296.0 * (channels[i].hiLIM - channels[i].loLIM);
                ELSE
                    channels[i].outputValue := channels[i].loLIM
                        + raw / 27648.0 * (channels[i].hiLIM - channels[i].loLIM);
                END_IF;
            ELSIF channels[i].measuringMode = 1 THEN
                channels[i].outputValue := raw / 10.0;
            ELSE
                channels[i].outputValue := raw / 100.0;
            END_IF;
        END_IF;
    END_IF;
END_FOR;

(* ---- M02_mode_check_off.st ---- *)
TYPE ST_AnalogChannel :
STRUCT
    enable        : BOOL;
    hiLIM         : REAL;
    loLIM         : REAL;
    bipolar       : BOOL;
    measuringMode : INT;
    retVal        : WORD;
    outputValue   : REAL;
END_STRUCT
END_TYPE

(* Q08 Analog Batch Processing - reference solution.
   The task declares ARRAY[*]; this reference fixes the length at 2 so that it
   can be compiled and exercised by the test harness. *)
FUNCTION_BLOCK FB_Q08
VAR_INPUT
    count : DINT;
END_VAR
VAR_IN_OUT
    analogValues : ARRAY[1..2] OF INT;
    channels     : ARRAY[1..2] OF ST_AnalogChannel;
END_VAR
VAR
    i   : DINT;
    raw : REAL;
END_VAR

FOR i := 1 TO 2 DO
    IF i <= count AND channels[i].enable THEN
        IF FALSE THEN
            channels[i].retVal := 16#8001;
        ELSIF channels[i].hiLIM <= channels[i].loLIM THEN
            channels[i].retVal := 16#8002;
        ELSE
            channels[i].retVal := 16#0000;
            raw := INT_TO_REAL(analogValues[i]);
            IF channels[i].measuringMode = 0 THEN
                IF channels[i].bipolar THEN
                    channels[i].outputValue := channels[i].loLIM
                        + (raw + 27648.0) / 55296.0 * (channels[i].hiLIM - channels[i].loLIM);
                ELSE
                    channels[i].outputValue := channels[i].loLIM
                        + raw / 27648.0 * (channels[i].hiLIM - channels[i].loLIM);
                END_IF;
            ELSIF channels[i].measuringMode = 1 THEN
                channels[i].outputValue := raw / 10.0;
            ELSE
                channels[i].outputValue := raw / 100.0;
            END_IF;
        END_IF;
    END_IF;
END_FOR;

(* ---- M03_no_window_check.st ---- *)
(* Q09 Calculate Moving Average - reference solution *)
FUNCTION_BLOCK FB_Q09
VAR_INPUT
    cyclicExecution : BOOL;
    trigger         : BOOL;
    value           : LREAL;
    windowSize      : INT;
    reset           : BOOL;
END_VAR
VAR_OUTPUT
    average            : LREAL;
    windowSizeReached  : BOOL;
    error              : BOOL;
    status             : WORD;
END_VAR
VAR
    buf   : ARRAY[0..99] OF LREAL;
    count : INT;
    head  : INT;
    sum   : LREAL;
    prevTrig : BOOL;
    doRead : BOOL;
    i : INT;
END_VAR

IF FALSE THEN
    error := TRUE;
    status := 16#8200;
    average := 0;
    windowSizeReached := FALSE;
    prevTrig := trigger;
    RETURN;
END_IF;
error := FALSE;
status := 16#0000;

IF reset THEN
    count := 0;
    head := 0;
    sum := 0;
    average := 0;
    windowSizeReached := FALSE;
    prevTrig := trigger;
    RETURN;
END_IF;

IF cyclicExecution THEN
    doRead := TRUE;
ELSE
    doRead := trigger AND NOT prevTrig;
END_IF;
prevTrig := trigger;

IF doRead THEN
    IF count < windowSize THEN
        buf[head] := value;
        sum := sum + value;
        count := count + 1;
    ELSE
        sum := sum - buf[head];
        buf[head] := value;
        sum := sum + value;
    END_IF;
    head := head + 1;
    IF head >= windowSize THEN
        head := 0;
    END_IF;
END_IF;

IF count > 0 THEN
    average := sum / INT_TO_LREAL(count);
ELSE
    average := 0;
END_IF;
windowSizeReached := count >= windowSize;

(* ---- M03_trigger_level.st ---- *)
(* Q09 Calculate Moving Average - reference solution *)
FUNCTION_BLOCK FB_Q09
VAR_INPUT
    cyclicExecution : BOOL;
    trigger         : BOOL;
    value           : LREAL;
    windowSize      : INT;
    reset           : BOOL;
END_VAR
VAR_OUTPUT
    average            : LREAL;
    windowSizeReached  : BOOL;
    error              : BOOL;
    status             : WORD;
END_VAR
VAR
    buf   : ARRAY[0..99] OF LREAL;
    count : INT;
    head  : INT;
    sum   : LREAL;
    prevTrig : BOOL;
    doRead : BOOL;
    i : INT;
END_VAR

IF windowSize < 1 OR windowSize > 100 THEN
    error := TRUE;
    status := 16#8200;
    average := 0;
    windowSizeReached := FALSE;
    prevTrig := trigger;
    RETURN;
END_IF;
error := FALSE;
status := 16#0000;

IF reset THEN
    count := 0;
    head := 0;
    sum := 0;
    average := 0;
    windowSizeReached := FALSE;
    prevTrig := trigger;
    RETURN;
END_IF;

IF cyclicExecution THEN
    doRead := TRUE;
ELSE
    doRead := trigger;
END_IF;
prevTrig := trigger;

IF doRead THEN
    IF count < windowSize THEN
        buf[head] := value;
        sum := sum + value;
        count := count + 1;
    ELSE
        sum := sum - buf[head];
        buf[head] := value;
        sum := sum + value;
    END_IF;
    head := head + 1;
    IF head >= windowSize THEN
        head := 0;
    END_IF;
END_IF;

IF count > 0 THEN
    average := sum / INT_TO_LREAL(count);
ELSE
    average := 0;
END_IF;
windowSizeReached := count >= windowSize;

(* ---- M04_no_fault.st ---- *)
(* Q10 Temperature Logic Control - reference solution *)
FUNCTION_BLOCK FB_Q10
VAR_INPUT
    TemperatureSensorInput : REAL;
    SetTemperature         : REAL;
END_VAR
VAR_OUTPUT
    CurrentTemperature : REAL;
    SetTempDisplay     : REAL;
    HeaterStatus       : BOOL;
    OverheatProtection : BOOL;
    HeaterOutput       : BOOL;
END_VAR
VAR
    runTimer  : TON;
    coolTimer : TON;
    sensorFault : BOOL;
END_VAR

CurrentTemperature := TemperatureSensorInput;
SetTempDisplay := SetTemperature;
sensorFault := FALSE;

runTimer(IN := HeaterOutput, PT := T#5S);
IF runTimer.Q THEN
    OverheatProtection := TRUE;
END_IF;

coolTimer(IN := OverheatProtection, PT := T#3S);
IF coolTimer.Q THEN
    OverheatProtection := FALSE;
END_IF;

IF sensorFault OR OverheatProtection THEN
    HeaterOutput := FALSE;
ELSIF TemperatureSensorInput < SetTemperature THEN
    HeaterOutput := TRUE;
ELSE
    HeaterOutput := FALSE;
END_IF;

HeaterStatus := HeaterOutput;

(* ---- M04_no_overheat.st ---- *)
(* Q10 Temperature Logic Control - reference solution *)
FUNCTION_BLOCK FB_Q10
VAR_INPUT
    TemperatureSensorInput : REAL;
    SetTemperature         : REAL;
END_VAR
VAR_OUTPUT
    CurrentTemperature : REAL;
    SetTempDisplay     : REAL;
    HeaterStatus       : BOOL;
    OverheatProtection : BOOL;
    HeaterOutput       : BOOL;
END_VAR
VAR
    runTimer  : TON;
    coolTimer : TON;
    sensorFault : BOOL;
END_VAR

CurrentTemperature := TemperatureSensorInput;
SetTempDisplay := SetTemperature;
sensorFault := TemperatureSensorInput < 0.0 OR TemperatureSensorInput > 100.0;

runTimer(IN := HeaterOutput, PT := T#5S);
(* no overheat *)

coolTimer(IN := OverheatProtection, PT := T#3S);
IF coolTimer.Q THEN
    OverheatProtection := FALSE;
END_IF;

IF sensorFault OR OverheatProtection THEN
    HeaterOutput := FALSE;
ELSIF TemperatureSensorInput < SetTemperature THEN
    HeaterOutput := TRUE;
ELSE
    HeaterOutput := FALSE;
END_IF;

HeaterStatus := HeaterOutput;

(* ---- M05_button_level.st ---- *)
FUNCTION_BLOCK M05_ProdLine
VAR_INPUT
    Mode : BOOL;
    ForwardButton : BOOL;
    ReverseButton : BOOL;
    SensorA : BOOL;
    SensorB : BOOL;
    SensorC : BOOL;
    ButtonA : BOOL;
    ButtonB : BOOL;
    ButtonC : BOOL;
END_VAR
VAR_OUTPUT
    MotorForward : BOOL;
    MotorReverse : BOOL;
    CompletionLight : BOOL;
END_VAR
VAR
    step : INT;   (* 0=at A waiting 1=A->B 2=at B waiting 3=B->C 4=at C done *)
    prevA : BOOL;
    prevB : BOOL;
    prevC : BOOL;
END_VAR

IF NOT Mode THEN
    (* manual mode with forward/reverse interlock *)
    MotorForward := ForwardButton AND NOT ReverseButton;
    MotorReverse := ReverseButton AND NOT ForwardButton;
    CompletionLight := FALSE;
ELSE
    MotorReverse := FALSE;
    IF step = 0 THEN
        MotorForward := FALSE;
        IF SensorA AND ButtonA THEN
            step := 1;
        END_IF;
    ELSIF step = 1 THEN
        MotorForward := TRUE;
        IF SensorB THEN
            MotorForward := FALSE;
            step := 2;
        END_IF;
    ELSIF step = 2 THEN
        MotorForward := FALSE;
        IF ButtonB THEN
            step := 3;
        END_IF;
    ELSIF step = 3 THEN
        MotorForward := TRUE;
        IF SensorC THEN
            MotorForward := FALSE;
            step := 4;
        END_IF;
    ELSE
        (* step 4: at C *)
        MotorForward := FALSE;
        IF ButtonC THEN
            CompletionLight := TRUE;
        END_IF;
        IF NOT SensorC THEN
            CompletionLight := FALSE;
            step := 0;
        END_IF;
    END_IF;
END_IF;

prevA := ButtonA;
prevB := ButtonB;
prevC := ButtonC;

(* ---- M05_no_interlock.st ---- *)
FUNCTION_BLOCK M05_ProdLine
VAR_INPUT
    Mode : BOOL;
    ForwardButton : BOOL;
    ReverseButton : BOOL;
    SensorA : BOOL;
    SensorB : BOOL;
    SensorC : BOOL;
    ButtonA : BOOL;
    ButtonB : BOOL;
    ButtonC : BOOL;
END_VAR
VAR_OUTPUT
    MotorForward : BOOL;
    MotorReverse : BOOL;
    CompletionLight : BOOL;
END_VAR
VAR
    step : INT;   (* 0=at A waiting 1=A->B 2=at B waiting 3=B->C 4=at C done *)
    prevA : BOOL;
    prevB : BOOL;
    prevC : BOOL;
END_VAR

IF NOT Mode THEN
    (* manual mode with forward/reverse interlock *)
    MotorForward := ForwardButton;
    MotorReverse := ReverseButton;
    CompletionLight := FALSE;
ELSE
    MotorReverse := FALSE;
    IF step = 0 THEN
        MotorForward := FALSE;
        IF SensorA AND ButtonA AND NOT prevA THEN
            step := 1;
        END_IF;
    ELSIF step = 1 THEN
        MotorForward := TRUE;
        IF SensorB THEN
            MotorForward := FALSE;
            step := 2;
        END_IF;
    ELSIF step = 2 THEN
        MotorForward := FALSE;
        IF ButtonB AND NOT prevB THEN
            step := 3;
        END_IF;
    ELSIF step = 3 THEN
        MotorForward := TRUE;
        IF SensorC THEN
            MotorForward := FALSE;
            step := 4;
        END_IF;
    ELSE
        (* step 4: at C *)
        MotorForward := FALSE;
        IF ButtonC AND NOT prevC THEN
            CompletionLight := TRUE;
        END_IF;
        IF NOT SensorC THEN
            CompletionLight := FALSE;
            step := 0;
        END_IF;
    END_IF;
END_IF;

prevA := ButtonA;
prevB := ButtonB;
prevC := ButtonC;

(* ---- M06_count_level.st ---- *)
(* Q12 Slab Thickness Alarm and Fault History - reference solution
   Unit convention: CycleTime in ms, Slab_Runtime_Accumulator in ns (LTIME). *)
FUNCTION_BLOCK FB_Q12
VAR_INPUT
    THICKNESS_FAULT        : BOOL;
    THICKNESS_SIGNAL_VALID : BOOL;
    CUTTING_RUN            : BOOL;
    FaultTimestamp         : DINT;
    CycleTime              : TIME;
END_VAR
VAR_OUTPUT
    THICKNESS_ALARM          : BOOL;
    Slab_Fault_Counter       : UINT;
    Slab_Runtime_Accumulator : LTIME;
    Slab_Fault_History       : ARRAY[0..4] OF DINT;
END_VAR
VAR
    holdAcc  : UDINT;   (* ms *)
    accNs    : ULINT;   (* ns *)
    prevFlt  : BOOL;
    i        : INT;
END_VAR

IF NOT THICKNESS_SIGNAL_VALID THEN
    THICKNESS_ALARM := FALSE;
    holdAcc := 0;
    prevFlt := FALSE;
ELSE
    IF THICKNESS_FAULT THEN
        (* new fault: count and record *)
        Slab_Fault_Counter := Slab_Fault_Counter + 1;
        FOR i := 4 TO 1 BY -1 DO
            Slab_Fault_History[i] := Slab_Fault_History[i-1];
        END_FOR;
        Slab_Fault_History[0] := FaultTimestamp;
        THICKNESS_ALARM := TRUE;
        holdAcc := 0;
    END_IF;
    prevFlt := THICKNESS_FAULT;

    IF THICKNESS_ALARM THEN
        IF THICKNESS_FAULT THEN
            holdAcc := 0;                       (* hold while the fault persists *)
        ELSE
            holdAcc := holdAcc + TIME_TO_UDINT(CycleTime);
            IF holdAcc >= 500 THEN
                THICKNESS_ALARM := FALSE;
            END_IF;
        END_IF;
    END_IF;

    IF CUTTING_RUN AND NOT THICKNESS_FAULT THEN
        accNs := accNs + UDINT_TO_ULINT(TIME_TO_UDINT(CycleTime)) * 1000000;
        Slab_Runtime_Accumulator := ULINT_TO_LTIME(accNs);
    END_IF;
END_IF;

(* ---- M06_no_hold.st ---- *)
(* Q12 Slab Thickness Alarm and Fault History - reference solution
   Unit convention: CycleTime in ms, Slab_Runtime_Accumulator in ns (LTIME). *)
FUNCTION_BLOCK FB_Q12
VAR_INPUT
    THICKNESS_FAULT        : BOOL;
    THICKNESS_SIGNAL_VALID : BOOL;
    CUTTING_RUN            : BOOL;
    FaultTimestamp         : DINT;
    CycleTime              : TIME;
END_VAR
VAR_OUTPUT
    THICKNESS_ALARM          : BOOL;
    Slab_Fault_Counter       : UINT;
    Slab_Runtime_Accumulator : LTIME;
    Slab_Fault_History       : ARRAY[0..4] OF DINT;
END_VAR
VAR
    holdAcc  : UDINT;   (* ms *)
    accNs    : ULINT;   (* ns *)
    prevFlt  : BOOL;
    i        : INT;
END_VAR

IF NOT THICKNESS_SIGNAL_VALID THEN
    THICKNESS_ALARM := FALSE;
    holdAcc := 0;
    prevFlt := FALSE;
ELSE
    IF THICKNESS_FAULT AND NOT prevFlt THEN
        (* new fault: count and record *)
        Slab_Fault_Counter := Slab_Fault_Counter + 1;
        FOR i := 4 TO 1 BY -1 DO
            Slab_Fault_History[i] := Slab_Fault_History[i-1];
        END_FOR;
        Slab_Fault_History[0] := FaultTimestamp;
        THICKNESS_ALARM := TRUE;
        holdAcc := 0;
    END_IF;
    prevFlt := THICKNESS_FAULT;

    IF THICKNESS_ALARM THEN
        IF THICKNESS_FAULT THEN
            holdAcc := 0;                       (* hold while the fault persists *)
        ELSE
            holdAcc := holdAcc + TIME_TO_UDINT(CycleTime);
            THICKNESS_ALARM := FALSE;
        END_IF;
    END_IF;

    IF CUTTING_RUN AND NOT THICKNESS_FAULT THEN
        accNs := accNs + UDINT_TO_ULINT(TIME_TO_UDINT(CycleTime)) * 1000000;
        Slab_Runtime_Accumulator := ULINT_TO_LTIME(accNs);
    END_IF;
END_IF;

(* ---- M07_eco_everywhere.st ---- *)
(* Q13 Office HVAC Multi-mode Energy-Saving Control - reference solution *)
FUNCTION_BLOCK FB_Q13
VAR_INPUT
    OCCUPANCY_DETECTED : BOOL;
    ENERGY_SAVING_MODE : BOOL;
    HVAC_MODE_SELECTOR : INT;
END_VAR
VAR_OUTPUT
    SUPPLY_FAN_RUN       : BOOL;
    TEMP_SETPOINT_ADJUST : INT;
END_VAR
VAR
    startTimer : TON;
END_VAR

startTimer(IN := OCCUPANCY_DETECTED AND HVAC_MODE_SELECTOR <> 3, PT := T#30S);
SUPPLY_FAN_RUN := startTimer.Q;

IF HVAC_MODE_SELECTOR = 3 THEN
    TEMP_SETPOINT_ADJUST := 4;
ELSIF OCCUPANCY_DETECTED THEN
    TEMP_SETPOINT_ADJUST := 0;
ELSIF HVAC_MODE_SELECTOR = 1 THEN
    TEMP_SETPOINT_ADJUST := 2;
ELSIF HVAC_MODE_SELECTOR = 2 THEN
    TEMP_SETPOINT_ADJUST := 4;
ELSIF ENERGY_SAVING_MODE THEN
    TEMP_SETPOINT_ADJUST := 3;
ELSE
    TEMP_SETPOINT_ADJUST := 2;
END_IF;

(* ---- M07_no_delay.st ---- *)
(* Q13 Office HVAC Multi-mode Energy-Saving Control - reference solution *)
FUNCTION_BLOCK FB_Q13
VAR_INPUT
    OCCUPANCY_DETECTED : BOOL;
    ENERGY_SAVING_MODE : BOOL;
    HVAC_MODE_SELECTOR : INT;
END_VAR
VAR_OUTPUT
    SUPPLY_FAN_RUN       : BOOL;
    TEMP_SETPOINT_ADJUST : INT;
END_VAR
VAR
    startTimer : TON;
END_VAR

startTimer(IN := OCCUPANCY_DETECTED AND HVAC_MODE_SELECTOR <> 3, PT := T#30S);
SUPPLY_FAN_RUN := OCCUPANCY_DETECTED AND HVAC_MODE_SELECTOR <> 3;

IF HVAC_MODE_SELECTOR = 3 THEN
    TEMP_SETPOINT_ADJUST := 4;
ELSIF OCCUPANCY_DETECTED THEN
    TEMP_SETPOINT_ADJUST := 0;
ELSIF HVAC_MODE_SELECTOR = 1 THEN
    TEMP_SETPOINT_ADJUST := 1;
ELSIF HVAC_MODE_SELECTOR = 2 THEN
    TEMP_SETPOINT_ADJUST := 4;
ELSIF ENERGY_SAVING_MODE THEN
    TEMP_SETPOINT_ADJUST := 3;
ELSE
    TEMP_SETPOINT_ADJUST := 2;
END_IF;

(* ---- M08_no_segcount.st ---- *)
(* Q14 IPv4 Parsing with Format and Range Checks - reference solution *)
FUNCTION_BLOCK FB_Q14
VAR_INPUT
    ipText : STRING(254);
END_VAR
VAR_OUTPUT
    ipValue : UDINT;
END_VAR
VAR
    i, n, segCount, digits, segVal : INT;
    ch : BYTE;
    acc : UDINT;
    ok : BOOL;
    pText : POINTER TO BYTE;
END_VAR

ipValue := 0;
acc := 0;
segCount := 0;
digits := 0;
segVal := 0;
ok := TRUE;
pText := ADR(ipText);
n := 0;
WHILE n < 254 AND pText[n] <> 0 DO
    n := n + 1;
END_WHILE;

IF n = 0 THEN
    RETURN;
END_IF;

FOR i := 0 TO n - 1 DO
    ch := pText[i];
    IF ch >= 48 AND ch <= 57 THEN
        segVal := segVal * 10 + (BYTE_TO_INT(ch) - 48);
        digits := digits + 1;
        IF digits > 3 OR segVal > 255 THEN
            ok := FALSE;
        END_IF;
    ELSIF ch = 46 THEN
        IF digits = 0 THEN
            ok := FALSE;
        END_IF;
        acc := acc * 256 + INT_TO_UDINT(segVal);
        segCount := segCount + 1;
        segVal := 0;
        digits := 0;
        IF segCount > 3 THEN
            ok := FALSE;
        END_IF;
    ELSE
        ok := FALSE;
    END_IF;
END_FOR;

IF digits = 0 THEN
    ok := FALSE;
END_IF;
acc := acc * 256 + INT_TO_UDINT(segVal);
segCount := segCount + 1;

IF ok THEN
    ipValue := acc;
END_IF;

(* ---- M08_range_off.st ---- *)
(* Q14 IPv4 Parsing with Format and Range Checks - reference solution *)
FUNCTION_BLOCK FB_Q14
VAR_INPUT
    ipText : STRING(254);
END_VAR
VAR_OUTPUT
    ipValue : UDINT;
END_VAR
VAR
    i, n, segCount, digits, segVal : INT;
    ch : BYTE;
    acc : UDINT;
    ok : BOOL;
    pText : POINTER TO BYTE;
END_VAR

ipValue := 0;
acc := 0;
segCount := 0;
digits := 0;
segVal := 0;
ok := TRUE;
pText := ADR(ipText);
n := 0;
WHILE n < 254 AND pText[n] <> 0 DO
    n := n + 1;
END_WHILE;

IF n = 0 THEN
    RETURN;
END_IF;

FOR i := 0 TO n - 1 DO
    ch := pText[i];
    IF ch >= 48 AND ch <= 57 THEN
        segVal := segVal * 10 + (BYTE_TO_INT(ch) - 48);
        digits := digits + 1;
        IF digits > 3 OR segVal > 256 THEN
            ok := FALSE;
        END_IF;
    ELSIF ch = 46 THEN
        IF digits = 0 THEN
            ok := FALSE;
        END_IF;
        acc := acc * 256 + INT_TO_UDINT(segVal);
        segCount := segCount + 1;
        segVal := 0;
        digits := 0;
        IF segCount > 3 THEN
            ok := FALSE;
        END_IF;
    ELSE
        ok := FALSE;
    END_IF;
END_FOR;

IF digits = 0 THEN
    ok := FALSE;
END_IF;
acc := acc * 256 + INT_TO_UDINT(segVal);
segCount := segCount + 1;

IF ok AND segCount = 4 THEN
    ipValue := acc;
END_IF;
